Staubli VAL3: getTool.pgx

public program getTool(num x_nIndex, tool& x_tTool)
begin

  link(x_tTool,flange)
  x_tTool=tToolItem[x_nIndex].tTool

end
